{attribute 'linkalways'}
{attribute 'no_explicit_call' := 'Use the methods of this class'}
{attribute 'enable_dynamic_creation'}
FUNCTION_BLOCK DriveAxis_Simulated IMPLEMENTS I_DriveAxis
VAR
	notConnectedError : HardwareError := (isActive := TRUE, id := Constants.SIMULATOR_NOT_CONNECTED_ERROR_ID, text := 'Simulatoren er ikke tilkoblet');
	link : REFERENCE TO SimulatorLink;
	side : WheelSide;
	isEnabled : BOOL;
END_VAR

METHOD FB_init : BOOL
VAR_INPUT
	bInitRetains : BOOL;
	bInCopyCode : BOOL;
	simulator : REFERENCE TO SimulatorLink;
	mountedSide : WheelSide;
END_VAR
link REF= simulator;
side := mountedSide;
END_METHOD

METHOD Enable
isEnabled := TRUE;
WriteEnabled();
END_METHOD

METHOD Disable
isEnabled := FALSE;
SetVelocity(0);
WriteEnabled();
END_METHOD

METHOD SetVelocity
VAR_INPUT
	velocityInRadPerS : LREAL;
END_VAR
VAR
	limited : LREAL;
END_VAR
limited := LIMIT(-Parameters.maxWheelSpeedInRadPerS, velocityInRadPerS, Parameters.maxWheelSpeedInRadPerS);
IF NOT isEnabled THEN
	limited := 0;
END_IF
IF side = WheelSide.LEFT THEN
	SimulatorIo.command.leftWheelSetpointInRadPerS := limited;
ELSE
	SimulatorIo.command.rightWheelSetpointInRadPerS := limited;
END_IF
END_METHOD

METHOD TryReset : BOOL
TryReset := IsReady;
END_METHOD

METHOD PRIVATE WriteEnabled
IF side = WheelSide.LEFT THEN
	SimulatorIo.command.isLeftDriveEnabled := isEnabled;
ELSE
	SimulatorIo.command.isRightDriveEnabled := isEnabled;
END_IF
END_METHOD

PROPERTY PositionInRad : LREAL
GET
IF side = WheelSide.LEFT THEN
	PositionInRad := SimulatorIo.feedback.leftWheelAngleInRad;
ELSE
	PositionInRad := SimulatorIo.feedback.rightWheelAngleInRad;
END_IF
END_GET
END_PROPERTY

PROPERTY VelocityInRadPerS : LREAL
GET
IF side = WheelSide.LEFT THEN
	VelocityInRadPerS := SimulatorIo.feedback.leftWheelVelocityInRadPerS;
ELSE
	VelocityInRadPerS := SimulatorIo.feedback.rightWheelVelocityInRadPerS;
END_IF
END_GET
END_PROPERTY

PROPERTY IsReady : BOOL
GET
IsReady := __ISVALIDREF(link) AND_THEN link.IsConnected AND isEnabled;
END_GET
END_PROPERTY

PROPERTY Error : HardwareError
GET
IF NOT __ISVALIDREF(link) OR_ELSE NOT link.IsConnected THEN
	Error := notConnectedError;
END_IF
END_GET
END_PROPERTY

END_FUNCTION_BLOCK

(* stored: Version 1.1.0.1, ProductVersion 3.1.4026.12
   POU DriveAxis_Simulated: Id {41ea52d8-b4d0-5db6-81df-59cc5855790a}, SpecialFunc None
   Method FB_init: Id {a3b6b933-e68e-5617-8fbb-8315f0194dda}
   Method Enable: Id {ac4a18f5-de0c-5370-8a97-84bc61afc214}
   Method Disable: Id {f36ff31a-dcfd-53b4-acf4-1846e24a85dc}
   Method SetVelocity: Id {2685f0d0-0d34-5138-83cc-2c54b951dffa}
   Method TryReset: Id {a99ce1f4-6729-5dd1-a830-8f53d132fd66}
   Method WriteEnabled: Id {39a98399-0bbc-59ab-9d34-81a4657cb18c}
   Property PositionInRad: Id {d7612386-066b-5e66-bca6-fa15d574f5df}
   Get Get: Id {4e5639da-5722-5e75-beb0-ac257b3c733c}
   Property VelocityInRadPerS: Id {292cb838-070b-5e83-8a24-fea4e703ef3b}
   Get Get: Id {06957e18-d553-59e5-9a7d-99d9e4f339c1}
   Property IsReady: Id {3fac5cc4-92bb-5edc-a90a-0ba070ebda6b}
   Get Get: Id {29f57d54-8962-51f4-8096-dc991b5406a5}
   Property Error: Id {47dce12e-2656-5a0a-8e78-d407b36dde07}
   Get Get: Id {75a31627-176d-537c-a57c-5a8cd49f753a} *)
